# EPICS substitutions: iocs/motor/oriel-ioc/db/EMC18011.substitutions
# C's iocOriel EMC18011.substitutions row, P from st.cmd: controller
# motor 1 only, as C loads it. The controller only reports position when
# stopped, and only for the currently selected motor.
file "$(MOTOR)/db/motor.db"
{
pattern
{N,  M,        DTYP,        S,  DESC,          EGU,      DIR,  VELO,  VBAS,  ACCL,  BDST,  BVEL,  BACC,  MRES,  PREC,  DHLM,    DLLM,  INIT}
{1,  "m$(N)",  "EMC18011",  0,  "motor $(N)",  microns,  Pos,  10,    0.,    1.,    0,     1,     .2,    0.01,  3,     999999,  0.1,   ""}
}
